(* IEC 61131-3 sources: SortJet_MasterSPS_Aufbau.fbsproj/07_Auftragsverwaltung, 9 files *)

(* ---- Job.prg.st ---- *)
(* METADATA
{
	"v3Meta": {
		"objectGuid": "d795aefc-c30c-4a59-9340-fdd22ca20f71"
	}
}
*)
PROGRAM Job
VAR

  // BOOLEAN
  blMerkerMmiNichtOk        : BOOL;
  blMerkerNachrichtabsetzen : BOOL;
  blSendJobStatus           : BOOL;
  blTsSeiteFehlerGesetzt    : BOOL; // Fehler-Seite eines Transfershuttles in abpFehler gesetzt
  ablFehlerAktiv            : ARRAY[cERSTER_AUTOMATIKKREIS..cLETZTER_AUTOMATIKKREIS] OF BOOL;

  // WORD
  wlMinutenMmiNichtOk       : WORD;
  wlSekundenMmiNichtOk      : WORD;
  wlMilliSekundenMmiNichtOk : WORD;
  wlIndex                   : WORD := 0;
  wlSubIndex                : WORD := 0;
  wlFaecherwagen            : WORD := 0; // Ampel blau: Faecherwagenstation
  wlIndexAK                 : WORD := 0; // Ampel blau: Automatikkreis der Station (Index)
  wlAK                      : WORD := 0; // Ampel blau: Automatikkreis der Station
  wlIndexStationen          : WORD := 0;
  wIndexReset               : WORD := 0;
  wIndexCheck               : WORD := 0;
  wlIndexSeite              : WORD := 0; // Automatikkreis-Index der Seiten eines Transfershuttles

  // LREAL
  lrlAktuelleZeit : LREAL;
  lrlMmiNichtOk   : LREAL;

  // TIMER
  timelMmiNichtOk       : TIME;
  tonlNachrichtAbsetzen : TON;
  tonlMmiOk             : TON;

  // TRIGGER
  rtlMmiOk                  : R_TRIG;
  ftlMmiOk                  : F_TRIG;
  ftlNotHaltAusgeloest      : F_TRIG;
  rtlFehlerAutomatikkreis   : ARRAY[cERSTER_AUTOMATIKKREIS..cLETZTER_AUTOMATIKKREIS] OF R_TRIG;

  // Check Betriebsart
  i        : WORD;
  mask     : WORD;
  newValue : BOOL;
  oldValue : BOOL;

END_VAR
//-------------------------------------------------------------------------------------------------
// STOPPEN DES AUTOMATIK- BETRIEBS [NOT-AUS]
//-------------------------------------------------------------------------------------------------
(* Anmerkung:
   - Automatikkreise stoppen sollte Notaus
*)
IF ( NOT NotHalt.bpNotHaltOK AND NOT bgSicherheitstechnikBruecken )
   OR ( NOT bgMMIOK AND NOT bgMMIBruecken )
THEN
  FOR wlIndex := cERSTER_AUTOMATIKKREIS TO cLETZTER_AUTOMATIKKREIS DO
    M_Automatik_Aktiv[wlIndex]   := FALSE;
  END_FOR
  M_Automatik_Aktiv[cAUTOMATIKKREIS_TRANSFERSHUTTLE] := FALSE;

END_IF

FOR wlIndex := cERSTER_AUTOMATIKKREIS TO cLETZTER_AUTOMATIKKREIS DO
  tonAutomatik_Aktiv[wlIndex]( IN := M_Automatik_Aktiv[wlIndex] AND NOT Stop_Baustein.abpBetriebsstop[wlIndex], PT := t#1s );
END_FOR

//-------------------------------------------------------------------------------------------------
// AKTIONEN
//-------------------------------------------------------------------------------------------------
FehlerAktiv();
CheckBetriebsart();
Check_MMI_Verbindung();
SendBetriebsart();
SetHandfunktionen();
Job_Shuttle();
Job_Stationen();
Job_Fremdanlage();
Job_SystemCheck();
Job_Verfahrlogik();
Job_Speicherfachvalidierung();
Job_Faecherwagen();
AutomatikStop();
AutomatikStart();
StartCheck();
Hornsignal();
Ampelsignal();
AnzeigeIOs();
Zuweisung_Automatik();
END_PROGRAM

(* ---- Job_Faecherwagen.prg.st ---- *)
(* METADATA
{
	"v3Meta": {
		"objectGuid": "77979386-6e9b-45aa-8f8e-3d53a4bcfd74"
	}
}
*)
PROGRAM Job_Faecherwagen
VAR_INPUT

  // BOOL
  abpReset  : ARRAY [cERSTER_AUTOMATIKKREIS..cLETZTER_AUTOMATIKKREIS] OF BOOL;

END_VAR
VAR_OUTPUT

  // BOOLEAN
  abpFehler : ARRAY[cERSTER_AUTOMATIKKREIS..cLETZTER_AUTOMATIKKREIS] OF BOOL;

END_VAR
VAR

  // BOOL
  blErsterZyklus          : BOOL := TRUE;
  awMerkerStatusFaecherwagenstationen : ARRAY[0..29] OF WORD;

  // WORD
  wlIndex                    : WORD;
  wlIndexReset               : WORD;
  wlIndexFaecherwagenStation : WORD;

  // INT
  ilBitPosition              : INT;
  ilIndexWordArray           : INT;

  // DWORD
  dwDifference : DWORD;

  // TRIGGER
  rtlErwzungenesAuschleusen  : ARRAY [cERSTE_FAECHERWAGENSTATIONS_NR..cLETZTE_FAECHERWAGENSTATIONS_NR] OF R_TRIG;
  rtlErwzungenesEinschleusen : ARRAY [cERSTE_FAECHERWAGENSTATIONS_NR..cLETZTE_FAECHERWAGENSTATIONS_NR] OF R_TRIG;
  rtlFehler                  : ARRAY [cERSTE_FAECHERWAGENSTATIONS_NR..cLETZTE_FAECHERWAGENSTATIONS_NR] OF R_TRIG;
  rtlAutomatikKreis          : ARRAY [cERSTER_AUTOMATIKKREIS..cLETZTER_AUTOMATIKKREIS] OF R_TRIG;
  rtlSystemCheckKreis        : ARRAY [cERSTER_AUTOMATIKKREIS..cLETZTER_AUTOMATIKKREIS] OF R_TRIG;

  // ARRAY
  tonlUeberwachungFaecherwagenPosition  : ARRAY[cERSTE_FAECHERWAGENSTATIONS_NR..cLETZTE_FAECHERWAGENSTATIONS_NR] OF TON;
  rtlUeberwachungFaecherwagenPosition   : ARRAY[cERSTE_FAECHERWAGENSTATIONS_NR..cLETZTE_FAECHERWAGENSTATIONS_NR] OF R_TRIG;
  rtlUeberwachungFaecherwagenPosition2  : ARRAY[cERSTE_FAECHERWAGENSTATIONS_NR..cLETZTE_FAECHERWAGENSTATIONS_NR] OF R_TRIG;

END_VAR

VAR CONSTANT

  // WORD
  cBIT_ANZAHL_WORD : WORD := 16;

END_VAR

//-------------------------------------------------------------------------------------------------
// INITIALISIERUNG
//-------------------------------------------------------------------------------------------------
IF ( blErsterZyklus ) THEN
  blErsterZyklus := FALSE;
END_IF

//-------------------------------------------------------------------------------------------------
// BELADUNGS STATUS
//-------------------------------------------------------------------------------------------------
(* Hinweis:
   - Abfrage des Status der Faecherwagenstation
     => 0 = frei
     => 1 = belegt
   - Das MMI fragt an welche Beladestationen belegt sind. Steht in dem ersten Wort z.B. die 301 als SPS Nummer
     Steht im ersten Wort der Antwort der Status dieser Station (siehe nächste Nachricht)
*)
IF ( M_SB0_MMI_REQUESTSTATUSLOADINGSTATIONS OR SlowTask.rtrigECatOK.Q OR Job.rtlMmiOk.Q ) AND bgEtherCatOK THEN

  M_SB0_MMI_REQUESTSTATUSLOADINGSTATIONS := FALSE;

  (* Hinweis:
     - Werte zuruecksetzen
  *)
  wlIndex       := WORD#0;
  ilBitPosition := INT#0;

  (* Hinweis:
     - Der Index ist [MMI_Var] fix auf 0-29 angelegt
  *)
  FOR ilIndexWordArray := 0 TO 29 DO
    awSps2MmiStatusFaecherwagenstationen[ilIndexWordArray] := WORD#0;
  END_FOR

  (* Hinweis:
     - Status der Stationen wird Bit-Codiert uebergeben
       => z.B.: Bit 0 = 301 | Bit 15 = 316
  *)
  FOR wlIndexFaecherwagenStation := cERSTE_FAECHERWAGENSTATIONS_NR TO cLETZTE_FAECHERWAGENSTATIONS_NR DO

    (* Hinweis:
       - Ein Bit kann gesetzt als auch zurueck gesetzt werden
    *)
    IF aFaecherwagenstation[wlIndexFaecherwagenStation].bStatusStationInBeladePosition THEN
      awSps2MmiStatusFaecherwagenstationen[wlIndex] := BitToggleWord( IN := awSps2MmiStatusFaecherwagenstationen[wlIndex], POS := ilBitPosition );
    END_IF

    IF ( ilBitPosition >= ( WORD_TO_INT(cBIT_ANZAHL_WORD) - 1) ) THEN
      wlIndex := INT_TO_WORD(INCI( WORD_TO_INT(wlIndex), 30 ));
    END_IF

    ilBitPosition := INCI( ilBitPosition, WORD_TO_INT(cBIT_ANZAHL_WORD) );

  END_FOR

  MsgToMmi(auftragsnr_w := SB0_SPS_SETSTATUSLOADINGSTATIONS );

END_IF

(* Hinweis:
   - Status der Stationen erstellen
*)
wlIndex       := WORD#0;
ilBitPosition := INT#0;

FOR ilIndexWordArray := 0 TO 29 DO
  awMerkerStatusFaecherwagenstationen[ilIndexWordArray] := WORD#0;
END_FOR
FOR wlIndexFaecherwagenStation := cERSTE_FAECHERWAGENSTATIONS_NR TO cLETZTE_FAECHERWAGENSTATIONS_NR DO

  IF aFaecherwagenstation[wlIndexFaecherwagenStation].bStatusStationInBeladePosition THEN
    awMerkerStatusFaecherwagenstationen[wlIndex] := BitToggleWord( IN := awMerkerStatusFaecherwagenstationen[wlIndex], POS := ilBitPosition );
  END_IF

  IF ( ilBitPosition >= ( WORD_TO_INT(cBIT_ANZAHL_WORD) - 1) ) THEN
    wlIndex := INT_TO_WORD( INCI( WORD_TO_INT(wlIndex), 30 ));
  END_IF

  ilBitPosition := INCI( ilBitPosition, WORD_TO_INT(cBIT_ANZAHL_WORD) );

END_FOR

dwDifference := DINT_TO_DWORD(SysMemCmp( ADR ( awSps2MmiStatusFaecherwagenstationen ), ADR( awMerkerStatusFaecherwagenstationen ), SIZEOF( awMerkerStatusFaecherwagenstationen )));
IF( dwDifference <> 0 AND bgEtherCatOK ) THEN
  awSps2MmiStatusFaecherwagenstationen := awMerkerStatusFaecherwagenstationen;
  MsgToMmi(auftragsnr_w := SB0_SPS_SETSTATUSLOADINGSTATIONS );
END_IF

//-------------------------------------------------------------------------------------------------
// FEHLER DER FAECHERWAGENSTATIONEN
//-------------------------------------------------------------------------------------------------
(* Hinweis:
   - Ein Fehler der Station setzt den Fehler in ihren Automatikkreisen (wie bei Stationen und Shuttle),
     der Betriebsstop wertet abpFehler aus. Das Zuruecksetzen erfolgt in der Aktion Reset.
*)
FOR wlIndexFaecherwagenStation := cERSTE_FAECHERWAGENSTATIONS_NR TO cLETZTE_FAECHERWAGENSTATIONS_NR DO
  rtlFehler[wlIndexFaecherwagenStation]( CLK := starrFaecherwagenBasisParameter[wlIndexFaecherwagenStation].bFehler );
  IF ( rtlFehler[wlIndexFaecherwagenStation].Q ) THEN
    AutomatikFehlerSetzen( starrFaecherwagenBasisParameter[wlIndexFaecherwagenStation].stMKs.eaAutomatikkreis, abpFehler );
  END_IF
END_FOR
//-------------------------------------------------------------------------------------------------
// AKTIONEN
//-------------------------------------------------------------------------------------------------
FWAuftraege();
Reset();
END_PROGRAM

(* ---- Job_Fremdanlage.prg.st ---- *)
(* METADATA
{
	"v3Meta": {
		"objectGuid": "ac7cd821-755f-477f-9445-f7486c53354c"
	}
}
*)
PROGRAM Job_Fremdanlage
VAR_INPUT

  // BOOL
  abpReset                    : ARRAY[cAUTOMATIKKREIS_1..cLETZTER_AUTOMATIKKREIS] OF BOOL;

  // AUJFTRAGSSPEICHER
  AuftragsSpeicherFremdanlage : ARRAY [cERSTE_FREMDANLAGE_AUSLAUF..cLETZTE_FREMDANLAGE_EINLAUF] OF AuftragsSpeicherStationen;

  // AUFTRAGS-STRUKTUREN
  AuftragsdatenFremdanlage    : ARRAY [cERSTE_FREMDANLAGE_AUSLAUF..cLETZTE_FREMDANLAGE_EINLAUF]  OF Auftragsdaten_ST;

END_VAR
VAR_OUTPUT

  // BOOL
  abpFehler          : ARRAY [cERSTER_AUTOMATIKKREIS..cLETZTER_AUTOMATIKKREIS] OF BOOL;

END_VAR
VAR

  // BOOL
  blErsterZyklus               : BOOL := TRUE;
  blUeberwachungFolgeNachricht : BOOL := FALSE;
  ablNachrichtEmpfangen        : ARRAY [1..2] OF BOOL;

  // WORD
  wlIndex          : WORD := 0;
  wlIndexReset     : WORD := 0;

  // STRUCT
  stAuftragScheibenIDs   : Schnittstelle_ScheibenIDs;

  // STEPS
  astplEintransportFremdanlage  : ARRAY [cERSTE_FREMDANLAGE_AUSLAUF..cLETZTE_FREMDANLAGE_EINLAUF] OF Steps_TE;

END_VAR
VAR CONSTANT

  // BYTE
  cNACHRICHTEN_INDEX_1 : BYTE := 1;
  cNACHRICHTEN_INDEX_2 : BYTE := 2;

END_VAR
//-------------------------------------------------------------------------------------------------
// BAUSTEIN: INITIALISIERUNG
//-------------------------------------------------------------------------------------------------
IF ( blErsterZyklus ) THEN
  blErsterZyklus := FALSE;

  ablNachrichtEmpfangen[1]     := FALSE;
  ablNachrichtEmpfangen[2]     := FALSE;
  blUeberwachungFolgeNachricht := FALSE;

END_IF

//-------------------------------------------------------------------------------------------------
// BAUSTEIN: AUFTRAGSVERWALTUNG
//-------------------------------------------------------------------------------------------------
FOR wlIndex := cERSTE_FREMDANLAGE_AUSLAUF TO cLETZTE_FREMDANLAGE_EINLAUF DO

  AuftragsSpeicherFremdanlage[wlIndex]();

  IF AuftragsSpeicherFremdanlage[wlIndex].bpAuftragverfuegbar
     AND ( AuftragsdatenFremdanlage[wlIndex].wAuftrag = eStation_Kein_Auftrag
           OR AuftragsdatenFremdanlage[wlIndex].wAuftrag = eStation_Belegt
           OR AuftragsdatenFremdanlage[wlIndex].wAuftrag = eStation_Warte_Auf_Eintransport )
  THEN
    AuftragsSpeicherFremdanlage[wlIndex].bpNaechsterAuftrag := TRUE;
    AuftragsSpeicherFremdanlage[wlIndex]();
    AuftragsdatenFremdanlage[wlIndex] := AuftragsSpeicherFremdanlage[wlIndex].AktAuftrag;
  END_IF

END_FOR

//-------------------------------------------------------------------------------------------------
// AKTIONEN
//-------------------------------------------------------------------------------------------------
Reset();
Auftraege();

// Hinweis:
// - Auslauf- Fremdanlagen: Vorgaenger und Automatikkreis aus den MKs der Schnittstelle
FOR wlIndex := cERSTE_FREMDANLAGE_AUSLAUF TO cLETZTE_FREMDANLAGE_AUSLAUF DO

  IF __ISVALIDREF( starrFremdanlageAuslaufStationBasisParameter[wlIndex].stMKs ) THEN
    Fremdanlage( wFremdanlage                  := wlIndex,
                 wVorgaenger                   := starrFremdanlageAuslaufStationBasisParameter[wlIndex].stMKs.stSchnittstellendaten.wVorgaengerStation,
                 wAutomatikkreis               := TO_WORD( AutomatikkreisBestimmen( wlIndex ) ),
                 bDurchtransportierendeStation := FALSE );
  END_IF

END_FOR
END_PROGRAM

(* ---- Job_Shuttle.prg.st ---- *)
(* METADATA
{
	"v3Meta": {
		"objectGuid": "fdc13e48-e8ff-456a-879e-40351fd7e090"
	}
}
*)
PROGRAM Job_Shuttle
VAR_INPUT

  // BOOLEAN
  abpReset                              : ARRAY[cERSTER_AUTOMATIKKREIS..cLETZTER_AUTOMATIKKREIS]    OF BOOL;
  abpStarteParalleleBausteinAnsteuerung : ARRAY [cERSTES_TRANSFERSHUTTLE..cLETZTES_TRANSFERSHUTTLE] OF BOOL;
  abpSpeicherfachValidierung            : ARRAY [cERSTES_TRANSFERSHUTTLE..cLETZTES_TRANSFERSHUTTLE] OF BOOL;
  abpResetTransportkopplung             : ARRAY [cERSTES_TRANSFERSHUTTLE..cLETZTES_TRANSFERSHUTTLE] OF BOOL;

  // BAUSTEINE
  AuftragsSpeicherTransfershuttle  : ARRAY [cERSTES_TRANSFERSHUTTLE..cLETZTES_TRANSFERSHUTTLE]          OF AuftragsSpeicher;
  AuftragsSpeicherShuttle          : ARRAY [cERSTES_SHUTTLE..cLETZTES_SHUTTLE]                          OF AuftragsSpeicher;
  AuftragsSpeicherWand             : ARRAY [cERSTES_SHUTTLE..cLETZTES_SHUTTLE, cWAND_1..cANZAHL_WAENDE] OF AuftragsSpeicher;

  // STRUCT
  AuftragsdatenStation                       : ARRAY [cERSTES_SHUTTLE..cLETZTES_SHUTTLE]                                  OF Auftragsdaten_ST;
  AuftragsdatenWand                          : ARRAY [cERSTES_SHUTTLE..cLETZTES_SHUTTLE, cWAND_1..cANZAHL_WAENDE]         OF Auftragsdaten_ST;
  VorAbAuftragsDaten                         : ARRAY [cERSTES_SHUTTLE..cLETZTES_TRANSFERSHUTTLE, cWAND_1..cANZAHL_WAENDE] OF VorAbAuftragsdaten_ST; // Ermoeglicht ein paralleles abarbeiten von bestimmten Auftraegen
  VisuAuftragsdaten                          : ARRAY [cERSTES_SHUTTLE..cLETZTES_TRANSFERSHUTTLE]                          OF Visu_Auftraege_ST;
  AuftragsdatenTransfershuttle               : ARRAY [cERSTES_TRANSFERSHUTTLE..cLETZTES_TRANSFERSHUTTLE]                  OF Auftragsdaten_ST;
  starrAuftragsdatenSpeicherfachValidierung  : ARRAY [cERSTES_TRANSFERSHUTTLE..cLETZTES_TRANSFERSHUTTLE]                  OF Auftragsdaten_ST;

  LocalAuftragsSpeicher             : REFERENCE TO AuftragsSpeicher;

END_VAR
VAR_OUTPUT

  // BOOLEAN
  abpFehler : ARRAY[cERSTER_AUTOMATIKKREIS..cLETZTER_AUTOMATIKKREIS] OF BOOL;

END_VAR
VAR

  // BOOLEAN
  blErsterZyklus         : BOOL := TRUE;
  blFehler               : ARRAY [cERSTES_SHUTTLE..cLETZTES_SHUTTLE, cWAND_1..cANZAHL_WAENDE] OF BOOL;
  blFehlerTS             : ARRAY [cERSTES_TRANSFERSHUTTLE..cLETZTES_TRANSFERSHUTTLE] OF BOOL;

  // WORD
  wlIndex,
  wlIndexWand,
  wlIndexQuelle,
  wlIndexReset,
  wlLetzteScheibe,
  wlErsteScheibe                  : WORD;
  awlGlasSender                   : ARRAY [cERSTES_TRANSFERSHUTTLE..cLETZTES_TRANSFERSHUTTLE] OF WORD;
  awlVerbundTransfershuttle       : ARRAY [cERSTES_TRANSFERSHUTTLE..cLETZTES_TRANSFERSHUTTLE] OF WORD;
  awlStatusSpeichervalidierung    : ARRAY [cERSTES_TRANSFERSHUTTLE..cLETZTES_TRANSFERSHUTTLE] OF WORD;

  // TRIGGER
  rtlFehler   : ARRAY[cERSTES_SHUTTLE..cLETZTES_SHUTTLE, cWAND_1..cANZAHL_WAENDE] OF R_TRIG;
  rtlFehlerTS : ARRAY[cERSTES_TRANSFERSHUTTLE..cLETZTES_TRANSFERSHUTTLE] OF R_TRIG;

  // STEPS
  asteplSpeicherfachValidierung   : ARRAY [cERSTES_TRANSFERSHUTTLE..cLETZTES_TRANSFERSHUTTLE] OF Steps_TE;
  asteplFaecherwagenSuche         : ARRAY [cERSTES_SHUTTLE..cLETZTES_SHUTTLE] OF Steps_TE;

  // TON
  atonlWarteAufMasterAuftrag      : ARRAY [cERSTES_TRANSFERSHUTTLE..cLETZTES_TRANSFERSHUTTLE] OF TON;

  // SH - BAUSTEINE
  Querfahrt                       : ARRAY[cERSTES_SHUTTLE..cLETZTES_SHUTTLE] OF Shuttle_Querfahrt;
  Racksuche                       : ARRAY[cERSTES_SHUTTLE..cLETZTES_SHUTTLE] OF Shuttle_RackSuche;
  Eintransport                    : ARRAY[cERSTES_SHUTTLE..cLETZTES_SHUTTLE, cWAND_1..cANZAHL_WAENDE] OF Shuttle_Eintransport;
  Austransport                    : ARRAY[cERSTES_SHUTTLE..cLETZTES_SHUTTLE, cWAND_1..cANZAHL_WAENDE] OF Shuttle_Austransport;
  Durchtransport                  : ARRAY[cERSTES_SHUTTLE..cLETZTES_SHUTTLE, cWAND_1..cANZAHL_WAENDE] OF Shuttle_Durchtransport;
  VorabkomponentenAnsteuerung     : ARRAY[cERSTES_SHUTTLE..cLETZTES_SHUTTLE, cWAND_1..cANZAHL_WAENDE] OF Shuttle_Vorabkomponenten;

  // TS - BAUSTEINE
  TS_Querfahrt                    : ARRAY[cERSTES_TRANSFERSHUTTLE..cLETZTES_TRANSFERSHUTTLE] OF TS_Querfahrt;
  TS_Eintransport                 : ARRAY[cERSTES_TRANSFERSHUTTLE..cLETZTES_TRANSFERSHUTTLE] OF TS_Eintransport;
  TS_Austransport                 : ARRAY[cERSTES_TRANSFERSHUTTLE..cLETZTES_TRANSFERSHUTTLE] OF TS_Austransport;
  TS_Transportkopplung            : ARRAY[cERSTES_TRANSFERSHUTTLE..cLETZTES_TRANSFERSHUTTLE] OF TS_Transportkopplung;
  TS_Vortransport                 : ARRAY[cERSTES_TRANSFERSHUTTLE..cLETZTES_TRANSFERSHUTTLE] OF TS_Vortransport;

  wlAutomatikkreis2               : WORD := 2; // Variable mit dem Index zum Zugriff auf den 2. Automatikkreis Index. Benötigt zum Austricksen des Compilers

  Basis                           : REFERENCE TO StationBasisParameter_ST;

END_VAR

//-------------------------------------------------------------------------------------------------
// BAUSTEIN: INITIALISIERUNG
//-------------------------------------------------------------------------------------------------
IF ( blErsterZyklus ) THEN
  blErsterZyklus := FALSE;

  FOR wlIndex := cERSTES_SHUTTLE TO cLETZTES_SHUTTLE DO
    Querfahrt[wlIndex].wStation := wlIndex;
    Racksuche[wlIndex].wStation := wlIndex;
    FOR wlIndexWand := cWAND_1 TO cANZAHL_WAENDE DO
      Eintransport[wlIndex, wlIndexWand].wStation                := wlIndex;
      Eintransport[wlIndex, wlIndexWand].wWand                   := wlIndexWand;
      Austransport[wlIndex, wlIndexWand].wStation                := wlIndex;
      Austransport[wlIndex, wlIndexWand].wWand                   := wlIndexWand;
      VorabkomponentenAnsteuerung[wlIndex, wlIndexWand].wStation := wlIndex;
      VorabkomponentenAnsteuerung[wlIndex, wlIndexWand].wWand    := wlIndexWand;
    END_FOR
  END_FOR

END_IF

(* Hinweis [TRANSFERSHUTTLE]:
   - Transportkopplungen zurücksetzen, wenn vom Master-TS gefordert
*)
FOR wlIndex := cERSTES_TRANSFERSHUTTLE TO cLETZTES_TRANSFERSHUTTLE DO
  IF NOT starrTransfershuttleBasisParameter[wlIndex].stMKs.stStationsOptionen.stTransfershuttle.bMasterStation THEN
    IF abpResetTransportkopplung[wlIndex] THEN
      abpResetTransportkopplung[wlIndex] := FALSE;
      TS_Transportkopplung[wlIndex]( bpReset := TRUE );
      AuftragsdatenTransfershuttle[wlIndex].wAuftrag := eStation_Kein_Auftrag;
    END_IF
  END_IF
END_FOR

//-------------------------------------------------------------------------------------------------
// BAUSTEIN: AKTIONEN
//-------------------------------------------------------------------------------------------------
(* Hinweis:
   - Aufruf der Baustein-Aktionen
*)
Auftraege();

FOR wlIndex := cERSTES_SHUTTLE TO cLETZTES_SHUTTLE DO

  FOR wlIndexWand := cWAND_1 TO cANZAHL_WAENDE DO
    rtlFehler[wlIndex,wlIndexWand]( CLK := blFehler[wlIndex,wlIndexWand] );
    ShuttleWandAuftraege(wlIndex, wlIndexWand);
  END_FOR

  ShuttleQuerfahrt(wlIndex);

END_FOR

FOR wlIndex := cERSTES_TRANSFERSHUTTLE TO cLETZTES_TRANSFERSHUTTLE DO
  rtlFehlerTS[wlIndex]( CLK := blFehlerTS[wlIndex] );
  IF starrTransfershuttleBasisParameter[wlIndex].stMKs.stStationsOptionen.stTransfershuttle.bMasterStation THEN
    Master_Transfershuttle(wlIndex);
  ELSE
    Slave_Transfershuttle(wlIndex);
  END_IF
END_FOR

Reset();
Meldungen();
Verfahrfreigabe();

//-------------------------------------------------------------------------------------------------
// BAUSTEIN: AUFTRAGSVERWALTUNG
//-------------------------------------------------------------------------------------------------
(* Hinweis:
   - Die Auftraege mussen vor dem Aufruf der Steuerung abgehandelt werden [Grund: z.B: Vermeidung von Fehlern nach dem SystemCheck]
*)

// Auftragsdaten für das Shuttle, z.B. Querfahrt
FOR wlIndex := cERSTES_SHUTTLE TO cLETZTES_SHUTTLE DO

  AuftragsSpeicherShuttle[wlIndex]();

  IF ( AuftragsSpeicherShuttle[wlIndex].bpAuftragverfuegbar
       AND ( ( AuftragsdatenStation[wlIndex].wAuftrag = eStation_Kein_Auftrag )
             OR ( AuftragsdatenStation[wlIndex].wAuftrag = eStation_Belegt ) ) )
  THEN
    AuftragsSpeicherShuttle[wlIndex].bpNaechsterAuftrag := TRUE;
    AuftragsSpeicherShuttle[wlIndex]();
    AuftragsdatenStation[wlIndex] := AuftragsSpeicherShuttle[wlIndex].AktAuftrag;
  END_IF

END_FOR

// Auftragsdaten für die Shuttlewand, z.B. Eintransport
FOR wlIndex := cERSTES_SHUTTLE TO cLETZTES_SHUTTLE DO

  FOR wlIndexWand := cWAND_1 TO cANZAHL_WAENDE DO

    AuftragsSpeicherWand[wlIndex, wlIndexWand]();

    IF    AuftragsSpeicherWand[wlIndex, wlIndexWand].bpAuftragverfuegbar
          AND AuftragsdatenWand[wlIndex, wlIndexWand].wAuftrag = eStation_Kein_Auftrag
    THEN
      AuftragsSpeicherWand[wlIndex, wlIndexWand].bpNaechsterAuftrag := TRUE;
      AuftragsSpeicherWand[wlIndex, wlIndexWand]();
      AuftragsdatenWand[wlIndex, wlIndexWand] := AuftragsSpeicherWand[wlIndex, wlIndexWand].AktAuftrag ;
    END_IF

  END_FOR

END_FOR

// Auftragsdaten für das Transfershuttle
FOR wlIndex := cERSTES_TRANSFERSHUTTLE TO cLETZTES_TRANSFERSHUTTLE DO

  AuftragsSpeicherTransfershuttle[wlIndex]();

  IF ( AuftragsSpeicherTransfershuttle[wlIndex].bpAuftragverfuegbar
       AND AuftragsdatenTransfershuttle[wlIndex].wAuftrag = eStation_Kein_Auftrag )
  THEN
    AuftragsSpeicherTransfershuttle[wlIndex].bpNaechsterAuftrag := TRUE;
    AuftragsSpeicherTransfershuttle[wlIndex]();
    AuftragsdatenTransfershuttle[wlIndex] := AuftragsSpeicherTransfershuttle[wlIndex].AktAuftrag;
  END_IF

END_FOR
END_PROGRAM

(* ---- Job_Speicherfachvalidierung.prg.st ---- *)
(* METADATA
{
	"v3Meta": {
		"objectGuid": "98bc2d31-e6c9-4c6f-a95b-80ba3f2124c6"
	}
}
*)
PROGRAM Job_Speicherfachvalidierung
VAR

  // BOOL
  blTransfershuttleNummerPlausibel       : BOOL := FALSE;
  blTransfershuttleVerbundNichtPlausibel : BOOL := TRUE;

  // WORD
  wlStationsNummer : WORD;

END_VAR
//-------------------------------------------------------------------------------------------------
// BAUSTEIN: VALIDIERUNGSDATEN FUER DAS TRANSFERSHUTTLE
//-------------------------------------------------------------------------------------------------
(* Hinweis:
   - Gesondertere Pruefung mittels Transfershuttles da der Einlauf- Auslauf- Sensor (oder beide) belegt
      wurden und dies zu einem Stopp der Anlage gefuehrt hat. Das Fach wird nochmal ueberprüft bevor
      die Anlage wieder in den Automatikmodus versetzt werden kann.
*)
IF ( M_SB0_MMI_TRANSFERSHUTTLECHECK ) THEN
  M_SB0_MMI_TRANSFERSHUTTLECHECK := FALSE;

  blTransfershuttleNummerPlausibel :=  PruefungWertImIntervall ( wpWert:= tMmi2SpsInfo.wTransfershuttle_Nummer1,
                                                                 wpIntervallMin  := cERSTES_TRANSFERSHUTTLE,
                                                                 wpIntervallMax := cLETZTES_TRANSFERSHUTTLE );

  // Wenn die Station plausibel ist weiter, ansonsten Fehlermeldung ausgeben
  IF ( blTransfershuttleNummerPlausibel ) THEN

    // Prüfen ob der Speichervalidierung noch aktiv ist, wenn ja -> Fehlermeldung
    IF ( Job_Shuttle.abpSpeicherfachValidierung[tMmi2SpsInfo.wTransfershuttle_Nummer1] ) THEN
      wpgFehlerdaten[0] := tMmi2SpsInfo.wTransfershuttle_Nummer1;
      wpgFehlerdaten[1] := tMmi2SpsInfo.wTransfershuttle_Nummer1;
      SpsHinweis( eFehler_Station,
                  cMELDUNG_TS_SPEICHERVALIDIERUNG_NOCH_AKTIV,
                  tMmi2SpsInfo.wTransfershuttle_Nummer1,
                  AutomatikkreisBestimmen(tMmi2SpsInfo.wTransfershuttle_Nummer1),
                  wpgFehlerdaten );
    ELSE
      // ---------------------------------------------------------------------------------------
      //  PRUEFEN TRANSFERSHUTTLE VERBUND
      //
      //  Hinweis:
      //  - wTransfershuttle_Nummer2 = 0   => Vortransport mit nur einem Transfershuttle
      //  - wTransfershuttle_Nummer2 <> 0  => Vortransport im Transfershuttle-Verbund
      // ---------------------------------------------------------------------------------------

      IF ( tMmi2SpsInfo.wTransfershuttle_Nummer2 <> 0 ) THEN
        VailiderenTransfershuttleVerbund ( wTransferstation1 := tMmi2SpsInfo.wTransfershuttle_Nummer1 ,
                                           wTransferstation2 := tMmi2SpsInfo.wTransfershuttle_Nummer2 ,
                                           wTransferstationMaster => tMmi2SpsInfo.wTransfershuttle_Nummer1,
                                           wTransferstationSlave  => tMmi2SpsInfo.wTransfershuttle_Nummer2,
                                           bpFehler               => blTransfershuttleVerbundNichtPlausibel );
      END_IF

      wlStationsNummer := tMmi2SpsInfo.wTransfershuttle_Nummer1;

      Job_Shuttle.starrAuftragsdatenSpeicherfachValidierung[wlStationsNummer].wStationsNr           := tMmi2SpsInfo.wTransfershuttle_Nummer1;

      IF ( tMmi2SpsInfo.wTransfershuttle_GlasDicke = 0 ) THEN
        Job_Shuttle.starrAuftragsdatenSpeicherfachValidierung[wlStationsNummer].rAuftragsDicke      := 4.0;
      ELSE
        Job_Shuttle.starrAuftragsdatenSpeicherfachValidierung[wlStationsNummer].rAuftragsDicke      := 19.0;
      END_IF

      Job_Shuttle.starrAuftragsdatenSpeicherfachValidierung[wlStationsNummer].rStationsZielposition := tMmi2SpsInfo.rTransfershuttle_SollPosition1;
      Job_Shuttle.starrAuftragsdatenSpeicherfachValidierung[wlStationsNummer].wTransferstationsNr1  := 0;
      Job_Shuttle.starrAuftragsdatenSpeicherfachValidierung[wlStationsNummer].rTransferposition1    := 0;

      IF ( NOT blTransfershuttleVerbundNichtPlausibel ) THEN
        Job_Shuttle.starrAuftragsdatenSpeicherfachValidierung[wlStationsNummer].wTransferstationsNr2  := tMmi2SpsInfo.wTransfershuttle_Nummer2;
        Job_Shuttle.starrAuftragsdatenSpeicherfachValidierung[wlStationsNummer].rTransferposition2    := tMmi2SpsInfo.rTransfershuttle_SollPosition2;
      ELSE
        Job_Shuttle.starrAuftragsdatenSpeicherfachValidierung[wlStationsNummer].rTransferposition2    := 0;
        Job_Shuttle.starrAuftragsdatenSpeicherfachValidierung[wlStationsNummer].wTransferstationsNr2  := 0;
      END_IF

      Job_Shuttle.abpSpeicherfachValidierung[wlStationsNummer] := TRUE;
    END_IF

  ELSE
    wpgFehlerdaten[0] := tMmi2SpsInfo.wTransfershuttle_Nummer1;
    wpgFehlerdaten[1] := tMmi2SpsInfo.wTransfershuttle_Nummer1;
    SpsHinweis( eFehler_Station,
                cMELDUNG_AUFTRAGSDATEN_UNGUELTIGE_STATION,
                tMmi2SpsInfo.wTransfershuttle_Nummer1,
                AutomatikkreisBestimmen(tMmi2SpsInfo.wTransfershuttle_Nummer1),
                wpgFehlerdaten );

  END_IF

END_IF
END_PROGRAM

(* ---- Job_Stationen.prg.st ---- *)
(* METADATA
{
	"v3Meta": {
		"objectGuid": "9b3e7ff2-3a2c-4bce-8ea4-25f3e47febe0"
	}
}
*)
PROGRAM Job_Stationen
VAR_INPUT

  // BOOLEAN
  abpReset                              : ARRAY [cERSTER_AUTOMATIKKREIS..cLETZTER_AUTOMATIKKREIS] OF BOOL;
  abpAbbruchAnlegeauftrag               : ARRAY [cERSTE_STATION..cLETZTE_STATION] OF BOOL; // Hinweis: Wird ein Anlegeauftrag abgebrochen (M_SB0_MMI_SORTIERUNGCANCELQUEUEDATA) so darf die
  abpStarteParalleleBausteinAnsteuerung : ARRAY [cERSTE_STATION..cLETZTE_STATION, cWAND_1..cANZAHL_WAENDE] OF BOOL;
  abpResetTransportkopplung             : ARRAY [cERSTE_STATION..cLETZTE_STATION, cWAND_1..cANZAHL_WAENDE] OF BOOL;

  // AUJFTRAGSSPEICHER
  AuftragsSpeicherStation     : ARRAY [cERSTE_STATION..cLETZTE_STATION]                          OF AuftragsSpeicherStationen;
  AuftragsSpeicherWand        : ARRAY [cERSTE_STATION..cLETZTE_STATION, cWAND_1..cANZAHL_WAENDE] OF AuftragsSpeicherStationen;

  // AUFTRAGS-STRUKTUREN
  AuftragsdatenStation        : ARRAY [cERSTE_STATION..cLETZTE_STATION] OF Auftragsdaten_ST;
  AuftragsdatenWand           : ARRAY [cERSTE_STATION..cLETZTE_STATION, cWAND_1..cANZAHL_WAENDE] OF Auftragsdaten_ST;
  VisuAuftragsdaten           : ARRAY [cERSTE_STATION..cLETZTE_STATION] OF Visu_Auftraege_ST;

END_VAR
VAR_OUTPUT

  // BOOL
  abpFehler          : ARRAY [cERSTER_AUTOMATIKKREIS..cLETZTER_AUTOMATIKKREIS] OF BOOL;

END_VAR
VAR

  // BOOLEAN
  blErsterZyklus   : BOOL := TRUE;
  ablFreigabeZurParalleleBausteinAnsteuerung : ARRAY [cERSTE_STATION..cLETZTE_STATION, cWAND_1..cANZAHL_WAENDE] OF BOOL;
  ablMerkerLetzteScheibeStation              : ARRAY [cERSTE_STATION..cLETZTE_STATION, cWAND_1..cANZAHL_WAENDE] OF BOOL;
  ablFehler                                  : ARRAY [cERSTE_STATION..cLETZTE_STATION, cWAND_1..cANZAHL_WAENDE] OF BOOL;

  // WORD
  wlIndex,
  wlIndexWand,
  wlIndexReset,
  wlIndexAutoStart,
  wlLetzteScheibe,
  wlErsteScheibe : WORD;

  // INT
  ailScheibenZuQuittierenEintransport        : ARRAY [cERSTE_STATION..cLETZTE_STATION, cWAND_1..cANZAHL_WAENDE] OF INT; // Scheibenzaehlung fuer die Quittierung
  ailScheibenZuQuittierenAustransport        : ARRAY [cERSTE_STATION..cLETZTE_STATION, cWAND_1..cANZAHL_WAENDE] OF INT; // Scheibenzaehlung fuer die Quittierung

  // TRIGGER
  rtlFehler          : ARRAY[cERSTE_STATION..cLETZTE_STATION, cWAND_1..cANZAHL_WAENDE] OF R_TRIG;
  rtlStartAutomatik  : ARRAY[cERSTER_AUTOMATIKKREIS..cLETZTER_AUTOMATIKKREIS] OF R_TRIG;

  // BAUSTEINE
  Anlegen            : ARRAY[cERSTE_STATION..cLETZTE_STATION, cWAND_1..cANZAHL_WAENDE] OF Station_Anlegen;
  Abnehmen           : ARRAY[cERSTE_STATION..cLETZTE_STATION, cWAND_1..cANZAHL_WAENDE] OF Station_Abnehmen;
  Glashoehenmessung  : ARRAY[cERSTE_STATION..cLETZTE_STATION, cWAND_1..cANZAHL_WAENDE] OF Station_Glashoehenmessung;
  Glaslaengenmessung : ARRAY[cERSTE_STATION..cLETZTE_STATION, cWAND_1..cANZAHL_WAENDE] OF Station_Glaslaengenmessung;
  Eintransport       : ARRAY[cERSTE_STATION..cLETZTE_STATION, cWAND_1..cANZAHL_WAENDE] OF Station_Eintransport;
  Austransport       : ARRAY[cERSTE_STATION..cLETZTE_STATION, cWAND_1..cANZAHL_WAENDE] OF Station_Austransport;
  Durchtransport     : ARRAY[cERSTE_STATION..cLETZTE_STATION, cWAND_1..cANZAHL_WAENDE] OF Station_Durchtransport;
  Transportkopplung  : ARRAY[cERSTE_STATION..cLETZTE_STATION, cWAND_1..cANZAHL_WAENDE] OF Station_Transportkopplung;
  Messkopplung       : ARRAY[cERSTE_STATION..cLETZTE_STATION, cWAND_1..cANZAHL_WAENDE] OF Station_Messkopplung;
  Vortransport       : ARRAY[cERSTE_STATION..cLETZTE_STATION, cWAND_1..cANZAHL_WAENDE] OF Station_Vortransport;
  Querfahrt          : ARRAY[cERSTE_STATION..cLETZTE_STATION] OF Station_Querfahrt;

  // STRUCT
  stLokaleKopplungZielStation : REFERENCE TO StationBasisParameter_ST;
  stLokaleKopplungsStation    : REFERENCE TO StationBasisParameter_ST;

END_VAR
VAR CONSTANT

  // Stationen die nicht in den dynamischen Methoden aufgerufen werden dürfen
  awcAusgeschlosseneStationen : ARRAY[1..10] OF WORD := [ 218, 9(cSTATION_DEFAULT) ];

END_VAR
//-------------------------------------------------------------------------------------------------
// BAUSTEIN: INITIALISIERUNG
//-------------------------------------------------------------------------------------------------
IF blErsterZyklus THEN
  blErsterZyklus := FALSE;

END_IF

//-------------------------------------------------------------------------------------------------
// Transportkopplungen zurücksetzen, wenn vom Master gefordert
//-------------------------------------------------------------------------------------------------

FOR wlIndex := cERSTE_STATION TO cLETZTE_STATION DO
  FOR wlIndexWand := cWAND_1 TO cANZAHL_WAENDE DO
    IF abpResetTransportkopplung[wlIndex, wlIndexWand] THEN
      abpResetTransportkopplung[wlIndex, wlIndexWand] := FALSE;
      Transportkopplung[wlIndex, wlIndexWand]( bpReset := TRUE );
      Messkopplung[wlIndex, wlIndexWand]( bpReset := TRUE );
      AuftragsdatenWand[wlIndex, wlIndexWand].wAuftrag := eStation_Kein_Auftrag;
    END_IF
  END_FOR
END_FOR

//-------------------------------------------------------------------------------------------------
// BAUSTEIN: AKTIONEN
//-------------------------------------------------------------------------------------------------

Status_Automatikkreis_Start();

Auftraege();

Auftragsverwaltung();

Schnittstelle_Stationen();

FOR wlIndex := cERSTE_STATION TO cLETZTE_STATION DO
  FOR wlIndexWand := cWAND_1 TO cANZAHL_WAENDE DO
    rtlFehler[wlIndex, wlIndexWand]( CLK := ablFehler[wlIndex, wlIndexWand] );
    IF NOT findInWORDArray(awcAusgeschlosseneStationen, wlIndex) THEN
      Station(wlIndex, wlIndexWand);
    END_IF
  END_FOR
END_FOR

Reset();

Verfahrfreigabe();

Visu();
END_PROGRAM

(* ---- Job_SystemCheck.prg.st ---- *)
(* METADATA
{
	"v3Meta": {
		"objectGuid": "5553795f-6afb-4bc3-99ad-34d496c885e5"
	}
}
*)
PROGRAM Job_SystemCheck
VAR

  // WORD
  wlIndex   : WORD := 0;

END_VAR
//-------------------------------------------------------------------------------------------------
// AUFTRAEGE: SYSTEMCHECK STATUS STATION
//-------------------------------------------------------------------------------------------------
(* Hinweis:
   - Informationen ueber die Stationen
     => SystemCheck
*)
IF ( M_SB0_MMI_SYSTEMCHECKSTATION ) THEN
  M_SB0_MMI_SYSTEMCHECKSTATION := FALSE;

  CASE tMmi2SpsInfo.wSystemCheckStationMmiNummer OF

    cERSTES_TRANSFERSHUTTLE..cLETZTES_TRANSFERSHUTTLE: ;

      cERSTES_SHUTTLE..cLETZTES_SHUTTLE,
        cERSTE_STATION..cLETZTE_STATION:

      IF NOT ( PruefungWertImIntervall( wpWert:= tMmi2SpsInfo.wSystemCheckStationSlot, wpIntervallMin := cWAND_1, wpIntervallMax := cANZAHL_WAENDE )  ) THEN
        wpgFehlerdaten[0] := tMmi2SpsInfo.wSystemCheckStationMmiNummer;
        wpgFehlerdaten[1] := tMmi2SpsInfo.wSystemCheckStationSlot;
        SpsHinweis( eFehler_Station,
                    cMELDUNG_AUFTRAGSDATEN_UNGUELTIGE_WAND,
                    tMmi2SpsInfo.wSystemCheckStationMmiNummer,
                    AutomatikkreisBestimmen(tMmi2SpsInfo.wSystemCheckStationMmiNummer),
                    wpgFehlerdaten );

      ELSE

        abgDateStationCheck[tMmi2SpsInfo.wSystemCheckStationMmiNummer, tMmi2SpsInfo.wSystemCheckStationSlot].stAuftragsInformationen.wAuftragsInformationen := tMmi2SpsInfo.wSystemCheckStationTyp;
        abgDateStationCheck[tMmi2SpsInfo.wSystemCheckStationMmiNummer, tMmi2SpsInfo.wSystemCheckStationSlot].rStationsZielposition                          := tMmi2SpsInfo.rSystemCheckStationSollPosition;
        abgDateStationCheck[tMmi2SpsInfo.wSystemCheckStationMmiNummer, tMmi2SpsInfo.wSystemCheckStationSlot].wAnzahlScheiben                                := tMmi2SpsInfo.wSystemCheckStationScheibenanzahl;
        abgDateStationCheck[tMmi2SpsInfo.wSystemCheckStationMmiNummer, tMmi2SpsInfo.wSystemCheckStationSlot].rAuftragsLaenge                                := tMmi2SpsInfo.rSystemCheckStationScheibenlaenge;
        abgDateStationCheck[tMmi2SpsInfo.wSystemCheckStationMmiNummer, tMmi2SpsInfo.wSystemCheckStationSlot].wTransferstationsNr1                           := tMmi2SpsInfo.wSystemCheckStationZielstation;
        abgDateStationCheck[tMmi2SpsInfo.wSystemCheckStationMmiNummer, tMmi2SpsInfo.wSystemCheckStationSlot].bLetzteScheibe                                 := tMmi2SpsInfo.wSystemCheckStationLetzteScheibe.0;
        abgDateStationCheck[tMmi2SpsInfo.wSystemCheckStationMmiNummer, tMmi2SpsInfo.wSystemCheckStationSlot].wTransferwand                                  := tMmi2SpsInfo.wSystemCheckStationSlot;
        abgDateStationCheck[tMmi2SpsInfo.wSystemCheckStationMmiNummer, tMmi2SpsInfo.wSystemCheckStationSlot].rModellVersatzVorne                            := tMmi2SpsInfo.rSystemCheckModellVersatzVorne;
        abgDateStationCheck[tMmi2SpsInfo.wSystemCheckStationMmiNummer, tMmi2SpsInfo.wSystemCheckStationSlot].rModellVersatzHinten                           := tMmi2SpsInfo.rSystemCheckModellVersatzHinten;
        abgDateStationCheck[tMmi2SpsInfo.wSystemCheckStationMmiNummer, tMmi2SpsInfo.wSystemCheckStationSlot].bModell                                        := tMmi2SpsInfo.wSytstemCheckStationModellaktiv.0;
        abgDateStationCheck[tMmi2SpsInfo.wSystemCheckStationMmiNummer, tMmi2SpsInfo.wSystemCheckStationSlot].wBeschichtung                                  := tMmi2SpsInfo.wSystemCheckStationBeschichtungsSeite;
        abgDateStationCheck[tMmi2SpsInfo.wSystemCheckStationMmiNummer, tMmi2SpsInfo.wSystemCheckStationSlot].rAuftragsDicke                                 := WORD_TO_REAL(tMmi2SpsInfo.wSystemCheckScheibenDicke);
        abgDateStationCheck[tMmi2SpsInfo.wSystemCheckStationMmiNummer, tMmi2SpsInfo.wSystemCheckStationSlot].rAuftragsGewicht                               := tMmi2SpsInfo.rSystemcheckGlasGewicht;

        SystemCheck.abpStationsDatenErhalten[tMmi2SpsInfo.wSystemCheckStationMmiNummer, tMmi2SpsInfo.wSystemCheckStationSlot]  := TRUE;

      END_IF

    ELSE
      wpgFehlerdaten[0] := tMmi2SpsInfo.wSystemCheckStationMmiNummer;
      SpsHinweis( eFehler_Station,
                  cMELDUNG_SYSTEMCHECK_AUFTRAGSDATEN_UNGUELTIG,
                  tMmi2SpsInfo.wSystemCheckStationMmiNummer,
                  AutomatikkreisBestimmen(tMmi2SpsInfo.wSystemCheckStationMmiNummer),
                  wpgFehlerdaten );

  END_CASE

END_IF
END_PROGRAM

(* ---- Job_Verfahrlogik.prg.st ---- *)
(* METADATA
{
	"v3Meta": {
		"objectGuid": "e2245dfb-7a4f-4b2e-8ea2-abea4deaa4b5"
	}
}
*)
PROGRAM Job_Verfahrlogik
VAR
END_VAR

//-------------------------------------------------------------------------------------------------
// AUFTRAG: VERFAHRLOGIK [QUERFAHRT] SHUTTLE
//-------------------------------------------------------------------------------------------------
(* Hinweis:
   - Steuerung der Verfahrbewegungen durch die Oberflaeche
     => Verfahrlogik
*)
IF ( M_SB0_MMI_SHUTTLEVORABPOSITIONIERUNG ) THEN
  M_SB0_MMI_SHUTTLEVORABPOSITIONIERUNG := FALSE;

  CASE tMmi2SpsInfo.wVorabStationsNr OF

    cERSTE_STATION..cLETZTE_STATION:
      Job_Stationen.AuftragsSpeicherStation[tMmi2SpsInfo.wVorabStationsNr].NeuerAuftrag.rVorabPosition                    := tMmi2SpsInfo.rVorabPositionierung;
      Job_Stationen.AuftragsSpeicherStation[tMmi2SpsInfo.wVorabStationsNr].NeuerAuftrag.rVorabUpdateZeit                  := tMmi2SpsInfo.rVorabUpdateZeit;
      Job_Stationen.AuftragsSpeicherStation[tMmi2SpsInfo.wVorabStationsNr].NeuerAuftrag.rVorabBeschleunigung              := tMmi2SpsInfo.rVorabBeschleunigung;
      Job_Stationen.AuftragsSpeicherStation[tMmi2SpsInfo.wVorabStationsNr].NeuerAuftrag.rVorabBremsrampe                  := tMmi2SpsInfo.rVorabVerzoegern;
      Job_Stationen.AuftragsSpeicherStation[tMmi2SpsInfo.wVorabStationsNr].NeuerAuftrag.rVorabGeschwindigkeit             := tMmi2SpsInfo.rVorabGeschwindigkeit;
      Job_Stationen.AuftragsSpeicherStation[tMmi2SpsInfo.wVorabStationsNr].NeuerAuftrag.rNennstromBeschleunigungsphase    := tMmi2SpsInfo.rNennstromBeschleunigungsphase;
      Job_Stationen.AuftragsSpeicherStation[tMmi2SpsInfo.wVorabStationsNr].NeuerAuftrag.rNennstromKonstantfahrt           := tMmi2SpsInfo.rNennstromKonstantfahrt;
      Job_Stationen.AuftragsSpeicherStation[tMmi2SpsInfo.wVorabStationsNr].NeuerAuftrag.rZeitintervalBeschleunigungsphase := tMmi2SpsInfo.rZeitintervalBeschleunigungsphase;
      Job_Stationen.AuftragsSpeicherStation[tMmi2SpsInfo.wVorabStationsNr].NeuerAuftrag.wVorabAuftragstyp                 := tMmi2SpsInfo.wVorabAuftragstyp;

      Job_Stationen.AuftragsSpeicherStation[tMmi2SpsInfo.wVorabStationsNr].NeuerAuftrag.wAuftrag := eStation_Vorabpositionierung;
      Job_Stationen.AuftragsSpeicherStation[tMmi2SpsInfo.wVorabStationsNr](bpNeuerAuftrag := TRUE);

    cERSTES_TRANSFERSHUTTLE..cLETZTES_TRANSFERSHUTTLE:
      Job_Shuttle.AuftragsSpeicherTransfershuttle[tMmi2SpsInfo.wVorabStationsNr].NeuerAuftrag.rVorabPosition                    := tMmi2SpsInfo.rVorabPositionierung;
      Job_Shuttle.AuftragsSpeicherTransfershuttle[tMmi2SpsInfo.wVorabStationsNr].NeuerAuftrag.rVorabUpdateZeit                  := tMmi2SpsInfo.rVorabUpdateZeit;
      Job_Shuttle.AuftragsSpeicherTransfershuttle[tMmi2SpsInfo.wVorabStationsNr].NeuerAuftrag.rVorabBeschleunigung              := tMmi2SpsInfo.rVorabBeschleunigung;
      Job_Shuttle.AuftragsSpeicherTransfershuttle[tMmi2SpsInfo.wVorabStationsNr].NeuerAuftrag.rVorabBremsrampe                  := tMmi2SpsInfo.rVorabVerzoegern;
      Job_Shuttle.AuftragsSpeicherTransfershuttle[tMmi2SpsInfo.wVorabStationsNr].NeuerAuftrag.rVorabGeschwindigkeit             := tMmi2SpsInfo.rVorabGeschwindigkeit;
      Job_Shuttle.AuftragsSpeicherTransfershuttle[tMmi2SpsInfo.wVorabStationsNr].NeuerAuftrag.rNennstromBeschleunigungsphase    := tMmi2SpsInfo.rNennstromBeschleunigungsphase;
      Job_Shuttle.AuftragsSpeicherTransfershuttle[tMmi2SpsInfo.wVorabStationsNr].NeuerAuftrag.rNennstromKonstantfahrt           := tMmi2SpsInfo.rNennstromKonstantfahrt;
      Job_Shuttle.AuftragsSpeicherTransfershuttle[tMmi2SpsInfo.wVorabStationsNr].NeuerAuftrag.rZeitintervalBeschleunigungsphase := tMmi2SpsInfo.rZeitintervalBeschleunigungsphase;
      Job_Shuttle.AuftragsSpeicherTransfershuttle[tMmi2SpsInfo.wVorabStationsNr].NeuerAuftrag.wVorabAuftragstyp                 := tMmi2SpsInfo.wVorabAuftragstyp;

      Job_Shuttle.AuftragsSpeicherTransfershuttle[tMmi2SpsInfo.wVorabStationsNr].NeuerAuftrag.wAuftrag := eStation_Vorabpositionierung;
      Job_Shuttle.AuftragsSpeicherTransfershuttle[tMmi2SpsInfo.wVorabStationsNr](bpNeuerAuftrag := TRUE);

    cERSTES_SHUTTLE..cLETZTES_SHUTTLE:
      Job_Shuttle.AuftragsSpeicherShuttle[tMmi2SpsInfo.wVorabStationsNr].NeuerAuftrag.rVorabPosition                    := tMmi2SpsInfo.rVorabPositionierung;
      Job_Shuttle.AuftragsSpeicherShuttle[tMmi2SpsInfo.wVorabStationsNr].NeuerAuftrag.rVorabUpdateZeit                  := tMmi2SpsInfo.rVorabUpdateZeit;
      Job_Shuttle.AuftragsSpeicherShuttle[tMmi2SpsInfo.wVorabStationsNr].NeuerAuftrag.rVorabBeschleunigung              := tMmi2SpsInfo.rVorabBeschleunigung;
      Job_Shuttle.AuftragsSpeicherShuttle[tMmi2SpsInfo.wVorabStationsNr].NeuerAuftrag.rVorabBremsrampe                  := tMmi2SpsInfo.rVorabVerzoegern;
      Job_Shuttle.AuftragsSpeicherShuttle[tMmi2SpsInfo.wVorabStationsNr].NeuerAuftrag.rVorabGeschwindigkeit             := tMmi2SpsInfo.rVorabGeschwindigkeit;
      Job_Shuttle.AuftragsSpeicherShuttle[tMmi2SpsInfo.wVorabStationsNr].NeuerAuftrag.rNennstromBeschleunigungsphase    := tMmi2SpsInfo.rNennstromBeschleunigungsphase;
      Job_Shuttle.AuftragsSpeicherShuttle[tMmi2SpsInfo.wVorabStationsNr].NeuerAuftrag.rNennstromKonstantfahrt           := tMmi2SpsInfo.rNennstromKonstantfahrt;
      Job_Shuttle.AuftragsSpeicherShuttle[tMmi2SpsInfo.wVorabStationsNr].NeuerAuftrag.rZeitintervalBeschleunigungsphase := tMmi2SpsInfo.rZeitintervalBeschleunigungsphase;
      Job_Shuttle.AuftragsSpeicherShuttle[tMmi2SpsInfo.wVorabStationsNr].NeuerAuftrag.wVorabAuftragstyp                 := tMmi2SpsInfo.wVorabAuftragstyp;

      Job_Shuttle.AuftragsSpeicherShuttle[tMmi2SpsInfo.wVorabStationsNr].NeuerAuftrag.wAuftrag := eStation_Vorabpositionierung;
      Job_Shuttle.AuftragsSpeicherShuttle[tMmi2SpsInfo.wVorabStationsNr](bpNeuerAuftrag := TRUE);

    ELSE
      ;

  END_CASE

END_IF
END_PROGRAM

(* ---- SystemCheck.prg.st ---- *)
(* METADATA
{
	"v3Meta": {
		"objectGuid": "0b2e66de-e2de-4ed3-849b-e96a185ab44d"
	}
}
*)
PROGRAM SystemCheck
VAR_INPUT

  // BOOLEAN
  abpCheck                 : ARRAY [cERSTER_AUTOMATIKKREIS..cLETZTER_AUTOMATIKKREIS] OF BOOL;
  abpReset                 : ARRAY [cERSTER_AUTOMATIKKREIS..cLETZTER_AUTOMATIKKREIS] OF BOOL; // Fehler aus dem Resetbaustein heraus zurücksetzen
  abpStationsDatenErhalten : ARRAY [cERSTES_SHUTTLE..cLETZTE_STATION, cWAND_1..cANZAHL_WAENDE] OF BOOL;

END_VAR
VAR_OUTPUT

  // BOOL
  abpFehler        : ARRAY [cERSTER_AUTOMATIKKREIS..cLETZTER_AUTOMATIKKREIS] OF BOOL;

END_VAR
VAR

  // BOOL
  blErsterZyklus                      : BOOL := TRUE;
  ablTimeOutMeldungGenerieren         : ARRAY [cERSTER_AUTOMATIKKREIS..cLETZTER_AUTOMATIKKREIS] OF BOOL;
  ablStationFehlerImCheck             : ARRAY [cERSTER_AUTOMATIKKREIS..cLETZTER_AUTOMATIKKREIS] OF BOOL; // mind. eine Station hat den Check mit Fehler beendet
  blCheckAktiv                        : BOOL;
  ablCheck                            : ARRAY [cERSTER_AUTOMATIKKREIS..cLETZTER_AUTOMATIKKREIS, 1..cMAX_ANZAHL_SYSTEMCHECKZYKLEN] OF BOOL;
  ablCheckDone                        : ARRAY [cERSTER_AUTOMATIKKREIS..cLETZTER_AUTOMATIKKREIS, 1..cMAX_ANZAHL_SYSTEMCHECKZYKLEN] OF BOOL;
  ablStationCheckAktiv                : ARRAY[cERSTE_STATION..cLETZTE_STATION] OF BOOL;
  ablFWCheckAktiv                     : ARRAY[cERSTE_FAECHERWAGENSTATIONS_NR..cLETZTE_FAECHERWAGENSTATIONS_NR] OF BOOL;
  ablShuttleCheckAktiv                : ARRAY[cERSTES_SHUTTLE..cLETZTES_SHUTTLE] OF BOOL;

  // STEPS
  asteplCheck                         : ARRAY[cERSTER_AUTOMATIKKREIS..cLETZTER_AUTOMATIKKREIS, 1..cMAX_ANZAHL_SYSTEMCHECKZYKLEN] OF Steps_TE;

  // WORD
  wlIndex                            : WORD;
  wlIndexSystemcheckZyklus           : WORD;
  wlIndexAutomatikkreis              : WORD;
  wlIndexStationsnummer              : WORD;
  wlIndexQuitt                       : WORD;
  wlIndexQuittStation                : WORD;
  wlIndexQuittPartner                : WORD;
  wlAktiverZyklus                    : WORD;

  // REFERENCE
  stlQuittStation                    : REFERENCE TO StationBasisParameter_ST;

  // INT
  ailAnzahlStationenCheckAktiv       : ARRAY[cERSTER_AUTOMATIKKREIS..cLETZTER_AUTOMATIKKREIS] OF INT;
  ailAnzahlShuttleCheckAktiv         : ARRAY[cERSTER_AUTOMATIKKREIS..cLETZTER_AUTOMATIKKREIS] OF INT;
  ailAnzahlFWStationenCheckAktiv     : ARRAY[cERSTER_AUTOMATIKKREIS..cLETZTER_AUTOMATIKKREIS] OF INT;

  // TIMER
  atonlWarnungSystemCheckBeginnt     : ARRAY[cERSTER_AUTOMATIKKREIS..cLETZTER_AUTOMATIKKREIS] OF TON;
  atonlWaitCheck                     : ARRAY[cERSTER_AUTOMATIKKREIS..cLETZTER_AUTOMATIKKREIS] OF TON;
  atonlCheck                         : ARRAY[cERSTER_AUTOMATIKKREIS..cLETZTER_AUTOMATIKKREIS] OF TON;
  atonlCheckWarteAufMMIDaten         : ARRAY[cERSTER_AUTOMATIKKREIS..cLETZTER_AUTOMATIKKREIS] OF TON;
  tonlCheckAktiv                     : ton;

END_VAR
//-------------------------------------------------------------------------------------------------
// INITIALISIERUNG
//-------------------------------------------------------------------------------------------------
// Zeiger Initialisieren
//  - SystemCheck mit Vorgaenger- bzw. Nachfolger- Station
IF ( blErsterZyklus ) THEN
  blErsterZyklus := FALSE;

  FOR wlIndex := cERSTES_SHUTTLE TO cLETZTE_STATION DO
    abpStationsDatenErhalten[wlIndex,1] := FALSE;
  END_FOR

END_IF

// Check aktiv und Init nicht OK
blCheckAktiv := FALSE;
FOR wlIndex := cERSTER_AUTOMATIKKREIS TO cLETZTER_AUTOMATIKKREIS DO
  IF abpCheck[wlIndex] OR abpReset[wlIndex] THEN
    blCheckAktiv := TRUE;
  END_IF
END_FOR

Reset();
// Wenn kein Systemcheck aktiv -> Rausspringen
tonlCheckAktiv( IN  := NOT blCheckAktiv, PT := T#100MS);
IF tonlCheckAktiv.Q THEN
  RETURN; //Funktioniert noch nicht richtig
END_IF

//-------------------------------------------------------------------------------------------------
// TIMER
//-------------------------------------------------------------------------------------------------
(* Anmerkung:
   - Wartezeit bis mit dem SystemCheck begonnen wird
   - Die Sicherheitskreise müssen einen Moment lang quittiert sein, damit alle Antriebe hoch gelaufen sind

     SystemCheck starten
   - Verbindung zur MMI ist vorhanden
   - Freigabe [Rest ist nicht aktiv]
   - Sicherheitskreise geschlossen
   - Notaus nicht aktiv
   - Arbeitsdruck [Druckluft] ist in Ordnung
*)
FOR wlIndexAutomatikkreis := cERSTER_AUTOMATIKKREIS TO cLETZTER_AUTOMATIKKREIS DO

  atonlWaitCheck[wlIndexAutomatikkreis]( IN := ( M_INIT_OK
                                                 AND NotHalt.bpNotHaltOK
                                                 AND EtherCAT_Master.xConfigFinished
                                                 AND ( checkSafetyCircuitsClosedFromAutomaticCircuit(wlIndexAutomatikkreis, TRUE) OR bgSicherheitstechnikBruecken )
                                                 AND ( TCPMain.l_fb_SortjetHMI.o_b_WatchdogOk OR bgMMIBruecken )
                                                 AND StatusAnlage.bpAnlageOK ),
                                         PT := T#3S);

END_FOR

//-------------------------------------------------------------------------------------------------
// AKTIONEN
//-------------------------------------------------------------------------------------------------

Vorsteuerung();

FOR wlIndexAutomatikkreis := cERSTER_AUTOMATIKKREIS TO cLETZTER_AUTOMATIKKREIS DO
  FOR wlIndexSystemcheckZyklus := 1 TO wgAnzahlSystemcheckZyklen DO
    Systemcheck(wlIndexAutomatikkreis, wlIndexSystemcheckZyklus);
  END_FOR
END_FOR

Quittierung_Scheiben();
Meldungen();
END_PROGRAM
